// TIA Portal V21 export
// export: Created 2026-11-22T02:34:36.7967493Z, ExportSetting WithDefaults, DisplayName Totally Integrated Automation Portal, DisplayVersion V21 Update 3, DisplayName STEP 7 Professional, DisplayVersion V21 Update 3, DisplayName STEP 7 Safety, DisplayVersion V21, DisplayName Tech WebApplication, DisplayVersion V21, DisplayName WinCC Basic/Comfort/Advanced, DisplayVersion V21 Update 3, DisplayName WinCC Unified, DisplayVersion V21 Update 3
VBScript "SetS3"  Type=Sub
  SmartTags("D_State") = 3
  SmartTags("D_Bool") = True
  SmartTags("D_SInt") = 127
  SmartTags("D_Int") = 32767
  SmartTags("D_DInt") = 2147483647
  SmartTags("D_USInt") = 255
  SmartTags("D_UInt") = 65535
  SmartTags("D_UDInt") = 4294967295
  SmartTags("D_Real") = 123456.789
  SmartTags("D_LReal") = 1E+300
  SmartTags("D_String") = "Ünïcödé äöüß ÄÖÜ € – long text that is wider than the field 0123456789 ABCDEFGHIJ"
  SmartTags("D_DateTime") = DateSerial(2099, 12, 31) + TimeSerial(23, 59, 59)
  SmartTags("D_Pct") = 100
  SmartTags("D_Range") = 75
  SmartTags("D_Bits") = 4
  SmartTags("D_Vis") = True
  SmartTags("D_En") = False
  SmartTags("D_X") = 853
  SmartTags("D_Y") = 400
  SmartTags("D_Max") = 50
  SmartTags("D_Min") = -50
  SmartTags("D_TL") = 10
  SmartTags("D_BarR") = 5
